(* IEC 61131-3 sources: llm-plc-st-eval/codesys/dobles/B1, 5 files *)

(* ---- 01_Correcta.st ---- *)
(* DOBLE DE PRUEBA B1/Correcta - NO ES CORPUS. Esperado: veredicto 1 *)
FUNCTION_BLOCK FB_Motor
VAR_INPUT
    btnMarcha : BOOL;
    btnParo : BOOL;
    btnEmerg : BOOL;
END_VAR
VAR_OUTPUT
    motorOn : BOOL;
END_VAR
VAR
    bloqueo : BOOL;
END_VAR
IF btnEmerg THEN
    motorOn := FALSE;
    bloqueo := TRUE;
ELSE
    IF bloqueo AND NOT btnMarcha THEN
        bloqueo := FALSE;
    END_IF
    IF btnParo THEN
        motorOn := FALSE;
    ELSIF btnMarcha AND NOT bloqueo THEN
        motorOn := TRUE;
    END_IF
END_IF
END_FUNCTION_BLOCK

(* ---- 02_SinEnclavamiento.st ---- *)
(* DOBLE DE PRUEBA B1/SinEnclavamiento - NO ES CORPUS. Esperado: veredicto 2, falla en el paso 2 *)
FUNCTION_BLOCK FB_Motor
VAR_INPUT
    btnMarcha : BOOL;
    btnParo : BOOL;
    btnEmerg : BOOL;
END_VAR
VAR_OUTPUT
    motorOn : BOOL;
END_VAR
VAR
    nada : BOOL;
END_VAR
motorOn := btnMarcha AND NOT btnParo AND NOT btnEmerg;
END_FUNCTION_BLOCK

(* ---- 03_RearranqueTrasEmergencia.st ---- *)
(* DOBLE DE PRUEBA B1/RearranqueTrasEmergencia - NO ES CORPUS. Esperado: veredicto 2, falla en el paso 6 *)
FUNCTION_BLOCK FB_Motor
VAR_INPUT
    btnMarcha : BOOL;
    btnParo : BOOL;
    btnEmerg : BOOL;
END_VAR
VAR_OUTPUT
    motorOn : BOOL;
END_VAR
VAR
    nada : BOOL;
END_VAR
IF btnParo OR btnEmerg THEN
    motorOn := FALSE;
ELSIF btnMarcha THEN
    motorOn := TRUE;
END_IF
END_FUNCTION_BLOCK

(* ---- 04_EmergenciaNoDomina.st ---- *)
(* DOBLE DE PRUEBA B1/EmergenciaNoDomina - NO ES CORPUS. Esperado: veredicto 2, falla en el paso 5 *)
FUNCTION_BLOCK FB_Motor
VAR_INPUT
    btnMarcha : BOOL;
    btnParo : BOOL;
    btnEmerg : BOOL;
END_VAR
VAR_OUTPUT
    motorOn : BOOL;
END_VAR
VAR
    nada : BOOL;
END_VAR
IF btnMarcha THEN
    motorOn := TRUE;
ELSIF btnParo OR btnEmerg THEN
    motorOn := FALSE;
END_IF
END_FUNCTION_BLOCK

(* ---- 05_ParoInvertido.st ---- *)
(* DOBLE DE PRUEBA B1/ParoInvertido - NO ES CORPUS. Esperado: veredicto 2, falla en el paso 1 *)
FUNCTION_BLOCK FB_Motor
VAR_INPUT
    btnMarcha : BOOL;
    btnParo : BOOL;
    btnEmerg : BOOL;
END_VAR
VAR_OUTPUT
    motorOn : BOOL;
END_VAR
VAR
    nada : BOOL;
END_VAR
IF btnEmerg OR NOT btnParo THEN
    motorOn := FALSE;
ELSIF btnMarcha THEN
    motorOn := TRUE;
END_IF
END_FUNCTION_BLOCK
